KUKA KRL program: PrecProg.src

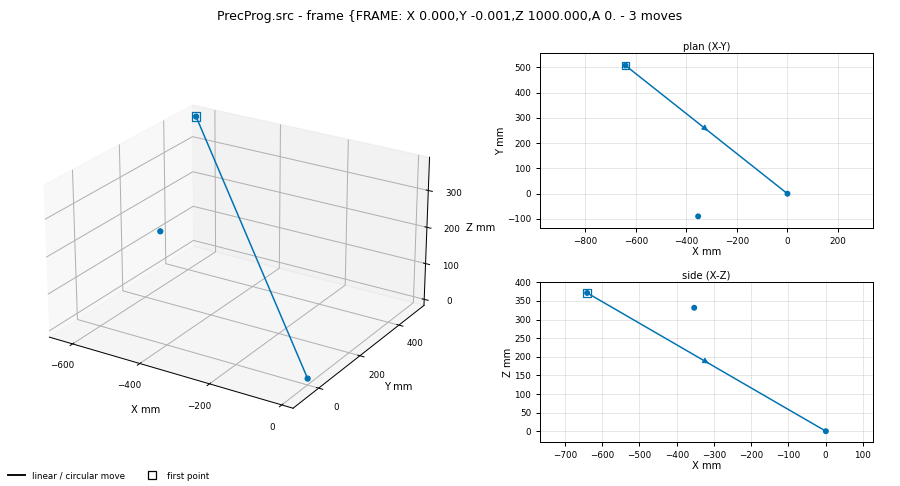
[picture p0: tool path of PrecProg.src in frame {FRAME: X 0.000,Y -0.001,Z 1000.000,A 0., 3 of 6 moves have a stored position in this frame; points joined in program order, loops and branches not executed]
&ACCESS RVP
&REL 1
&PARAM TEMPLATE = C:\KRC\Roboter\Template\vorgabe
&PARAM EDITMASK = *
DEF PrecProg ( )


; GLOBAL INTERRUPT DECL 3 WHEN $STOPMESS==TRUE DO IR_STOPM ( )
; INTERRUPT ON 3

;FOLD Initialise and set default speed
BAS (#INITMOV,0)
BAS (#VEL_PTP,100)
BAS (#ACC_PTP,20)
$VEL.CP=0.2
BAS (#TOOL,0)
BAS (#BASE,0)
;ENDFOLD

;;FOLD STARTPOS
;$BWDSTART = FALSE
;PDAT_ACT = PDEFAULT
;BAS(#PTP_DAT)
;FDAT_ACT = {TOOL_NO 0,BASE_NO 0,IPO_FRAME #BASE}
;BAS(#FRAMES)
;;ENDFOLD

$ADVANCE = 5

;FOLD ---- Quickly skip BCO ----
; PTP $AXIS_ACT
;ENDFOLD

;FOLD ---- GO HOME ----
; PTP {A1 0.000, A2 -90.000, A3 90.000, A4 0.000, A5 0.000, A6 0.000, E1 0, E2 0, E3 0, E4 0, E5 0, E6 0}
;ENDFOLD


; Program generated by RoboDK v6.0.7 for KUKA KR 10 R1440-2 on XX/XX/XXXX 18:00:00
; Using nominal kinematics.
; ---- Setting reference (Base) ----
$BASE = {FRAME: X 0.000,Y -0.001,Z 1000.000,A 0.123,B -0.500,C 90.000}
; --------------------------
; ---- Setting tool (TCP) ----
$TOOL = {FRAME: X 0.125,Y -0.375,Z 123.457,A 0.000,B 0.000,C -45.250}
; --------------------------
PTP {A1 12.34560,A2 -45.67890,A3 78.90130,A4 -0.50000,A5 0.49999,A6 180.00000}
LIN {X -640.585,Y 506.981,Z 371.534,A 150.000,B 50.000,C -165.500}
LIN {X 0.500,Y -0.500,Z 0.250,A 0.005,B -0.005,C 180.000}
PTP {A1 -12.34540,A2 45.67850,A3 -78.90000,A4 0.50000,A5 -0.00010,A6 -180.00000}
PTP {A1 -12.34540,A2 45.67850,A3 -78.90000,A4 0.50000,A5 -0.00010,A6 -180.00000}
$VEL.CP = 0.06667
WAIT SEC 0.002
WAIT SEC 1.000
LIN {X -353.026,Y -90.135,Z 331.702,A 178.023,B 40.650,C -169.444}
END
